// TIA Portal V21 export
VAR_GLOBAL   // PLC tag table "Standard-Variablentabelle"
   PositioningAxis_1_Actor_Interface_AddressIn AT %I266.0 : "PD_TEL105_IN";
   "PositioningAxis_1_Actor_Interface_AddressIn(1)" AT %I258.0 : "PD_TEL1_IN";
   PositioningAxis_1_Sensor1_Interface_AddressIn AT %I258.0 : "PD_TEL81_IN";
   "PositioningAxis_1_Actor_Interface_AddressIn(2)" AT %I258.0 : "PD_TEL105_IN";
   PositioningAxis_2_Actor_Interface_AddressIn AT %I280.0 : "PD_TEL105_IN";
   Einschubsachse_Actor_Interface_AddressIn AT %I12.0 : "PD_TEL3_IN";
   "Antrieb2_vertikale Achse_Actor_Interface_AddressIn" AT %I280.0 : "PD_TEL3_IN";
   "Antrieb2_vertikale Achse_Sensor1_Interface_AddressIn" AT %I280.0 : "PD_TEL103_IN";
   "Antrieb2_vertikale Achse_Actor_Interface_AddressIn(1)" AT %I280.0 : "PD_TEL1_IN";
   PositioningAxis_1_Actor_Interface_AddressOut AT %Q266.0 : "PD_TEL105_OUT";
   "PositioningAxis_1_Actor_Interface_AddressOut(1)" AT %Q258.0 : "PD_TEL1_OUT";
   PositioningAxis_1_Sensor1_Interface_AddressOut AT %Q258.0 : "PD_TEL81_OUT";
   "PositioningAxis_1_Actor_Interface_AddressOut(2)" AT %Q258.0 : "PD_TEL105_OUT";
   PositioningAxis_2_Actor_Interface_AddressOut AT %Q280.0 : "PD_TEL105_OUT";
   Einschubsachse_Actor_Interface_AddressOut AT %Q8.0 : "PD_TEL3_OUT";
   "Antrieb2_vertikale Achse_Actor_Interface_AddressOut" AT %Q280.0 : "PD_TEL3_OUT";
   "Antrieb2_vertikale Achse_Sensor1_Interface_AddressOut" AT %Q280.0 : "PD_TEL103_OUT";
   "Antrieb2_vertikale Achse_Actor_Interface_AddressOut(1)" AT %Q280.0 : "PD_TEL1_OUT";
   System_Byte AT %MB1 : Byte;
   FirstScan AT %M1.0 : Bool;
   DiagStatusUpdate AT %M1.1 : Bool;
   AlwaysTRUE AT %M1.2 : Bool;
   AlwaysFALSE AT %M1.3 : Bool;
   Clock_Byte AT %MB0 : Byte;
   Clock_10Hz AT %M0.0 : Bool;
   Clock_5Hz AT %M0.1 : Bool;
   "Clock_2.5Hz" AT %M0.2 : Bool;
   Clock_2Hz AT %M0.3 : Bool;
   "Clock_1.25Hz" AT %M0.4 : Bool;
   Clock_1Hz AT %M0.5 : Bool;
   "Clock_0.625Hz" AT %M0.6 : Bool;
   "Clock_0.5Hz" AT %M0.7 : Bool;
   state AT %MW50 : Int;
   Ventil_A AT %Q1.0 : Bool;
END_VAR
